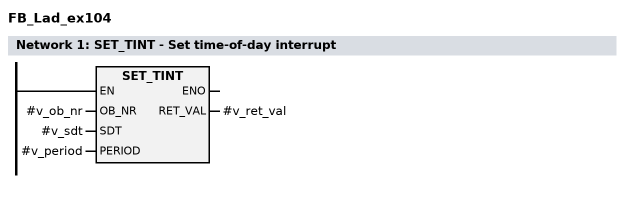
   #v_ret_val := SET_TINT(OB_NR := #v_ob_nr, SDT := #v_sdt, PERIOD := #v_period);
END_REGION
END_FUNCTION_BLOCK

FUNCTION_BLOCK "FB_Lad_ex105"   // FB30, LAD
{ S7_Optimized_Access := 'TRUE' }
   VAR_INPUT
      v_ob_nr : OB_Tod;
      v_sdt : DTL;
      v_local : Bool;
      v_period : Word;
      v_activate : Bool;
      v_ret_val : Int;
   END_VAR
BEGIN

REGION Network 1: SET_TINTL - Set time-of-day interrupt
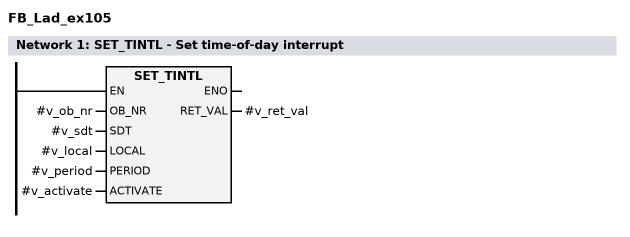
   #v_ret_val := SET_TINTL(OB_NR := #v_ob_nr,
                           SDT := #v_sdt,
                           LOCAL := #v_local,
                           PERIOD := #v_period,
                           ACTIVATE := #v_activate);
END_REGION
END_FUNCTION_BLOCK

FUNCTION_BLOCK "FB_Lad_ex106"   // FB31, LAD
{ S7_Optimized_Access := 'TRUE' }
   VAR_INPUT
      v_ob_nr : OB_Tod;
      v_ret_val : Int;
   END_VAR
BEGIN

REGION Network 1: CAN_TINT - Cancel time-of-day interrupt
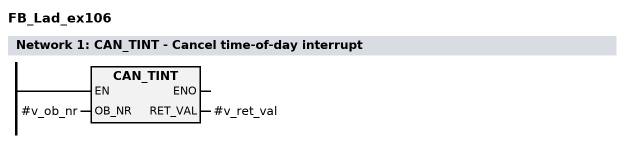
   #v_ret_val := CAN_TINT(OB_NR := #v_ob_nr);
END_REGION
END_FUNCTION_BLOCK

FUNCTION_BLOCK "FB_Lad_ex107"   // FB32, LAD
{ S7_Optimized_Access := 'TRUE' }
   VAR_INPUT
      v_ob_nr : OB_Tod;
      v_ret_val : Int;
   END_VAR
BEGIN

REGION Network 1: ACT_TINT - Enable time-of-day interrupt
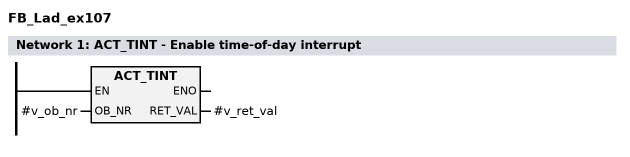
   #v_ret_val := ACT_TINT(OB_NR := #v_ob_nr);
END_REGION
END_FUNCTION_BLOCK

FUNCTION_BLOCK "FB_Lad_ex108"   // FB33, LAD
{ S7_Optimized_Access := 'TRUE' }
   VAR_INPUT
      v_ob_nr : OB_Tod;
      v_ret_val : Int;
   END_VAR
   VAR_OUTPUT
      v_status : Word;
   END_VAR
BEGIN

REGION Network 1: QRY_TINT - Query status of time-of-day interrupt
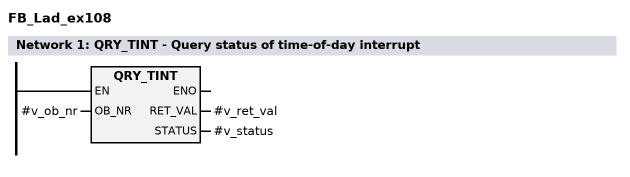
   #v_ret_val := QRY_TINT(OB_NR := #v_ob_nr, STATUS => #v_status);
END_REGION
END_FUNCTION_BLOCK

FUNCTION_BLOCK "FB_Lad_ex109"   // FB34, LAD
{ S7_Optimized_Access := 'TRUE' }
   VAR_INPUT
      v_ob_nr : Int;
      v_dtime : Time;
      v_sign : Word;
      v_ret_val : Int;
   END_VAR
BEGIN

REGION Network 1: SRT_DINT - Start time-delay interrupt
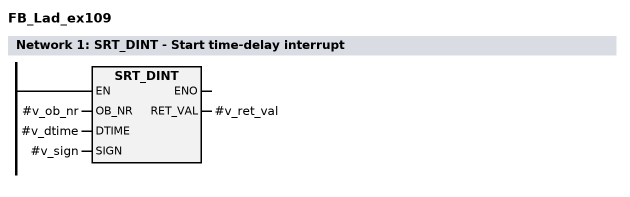
   #v_ret_val := SRT_DINT(OB_NR := #v_ob_nr, DTIME := #v_dtime, SIGN := #v_sign);
END_REGION
END_FUNCTION_BLOCK

FUNCTION_BLOCK "FB_Lad_ex110"   // FB35, LAD
{ S7_Optimized_Access := 'TRUE' }
   VAR_INPUT
      v_ob_nr : Int;
      v_ret_val : Int;
   END_VAR
BEGIN

REGION Network 1: CAN_DINT - Cancel time-delay interrupt
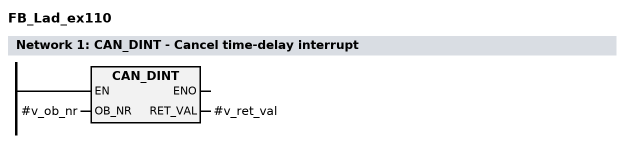
   #v_ret_val := CAN_DINT(OB_NR := #v_ob_nr);
END_REGION
END_FUNCTION_BLOCK

FUNCTION_BLOCK "FB_Lad_ex111"   // FB36, LAD
{ S7_Optimized_Access := 'TRUE' }
   VAR_INPUT
      v_ob_nr : Int;
      v_ret_val : Int;
   END_VAR
   VAR_OUTPUT
      v_status : Word;
   END_VAR
BEGIN

REGION Network 1: QRY_DINT - Query time-delay interrupt status
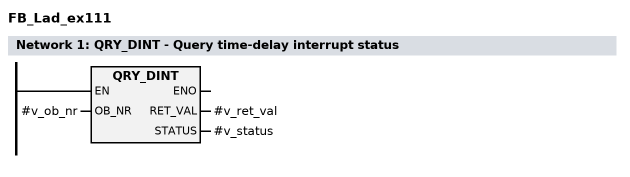
   #v_ret_val := QRY_DINT(OB_NR := #v_ob_nr, STATUS => #v_status);
END_REGION
END_FUNCTION_BLOCK

FUNCTION_BLOCK "FB_Lad_ex112"   // FB37, LAD
{ S7_Optimized_Access := 'TRUE' }
   VAR_INPUT
      v_prgflt_set_mask : DWord;
      v_accflt_set_mask : DWord;
      v_ret_val : Int;
   END_VAR
   VAR_OUTPUT
      v_prgflt_masked : DWord;
      v_accflt_masked : DWord;
   END_VAR
BEGIN

REGION Network 1: MSK_FLT - Mask synchronous error events
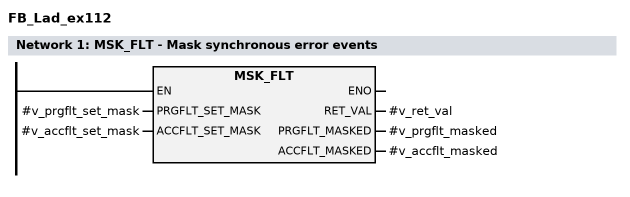
   #v_ret_val := MSK_FLT(PRGFLT_SET_MASK := #v_prgflt_set_mask,
                         ACCFLT_SET_MASK := #v_accflt_set_mask,
                         PRGFLT_MASKED => #v_prgflt_masked,
                         ACCFLT_MASKED => #v_accflt_masked);
END_REGION
END_FUNCTION_BLOCK

FUNCTION_BLOCK "FB_Lad_ex113"   // FB38, LAD
{ S7_Optimized_Access := 'TRUE' }
   VAR_INPUT
      v_prgflt_reset_mask : DWord;
      v_accflt_reset_mask : DWord;
      v_ret_val : Int;
   END_VAR
   VAR_OUTPUT
      v_prgflt_masked : DWord;
      v_accflt_masked : DWord;
   END_VAR
BEGIN

REGION Network 1: DMSK_FLT - Unmask synchronous error events
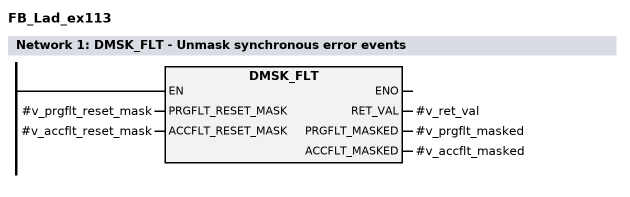
   #v_ret_val := DMSK_FLT(PRGFLT_RESET_MASK := #v_prgflt_reset_mask,
                          ACCFLT_RESET_MASK := #v_accflt_reset_mask,
                          PRGFLT_MASKED => #v_prgflt_masked,
                          ACCFLT_MASKED => #v_accflt_masked);
END_REGION
END_FUNCTION_BLOCK

FUNCTION_BLOCK "FB_Lad_ex114"   // FB39, LAD
{ S7_Optimized_Access := 'TRUE' }
   VAR_INPUT
      v_prgflt_query : DWord;
      v_accflt_query : DWord;
      v_ret_val : Int;
   END_VAR
   VAR_OUTPUT
      v_prgflt_clr : DWord;
      v_accflt_clr : DWord;
   END_VAR
BEGIN

REGION Network 1: READ_ERR - Read out event status register
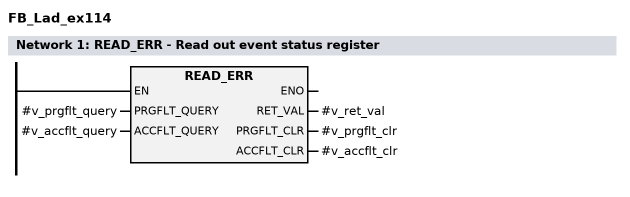
   #v_ret_val := READ_ERR(PRGFLT_QUERY := #v_prgflt_query,
                          ACCFLT_QUERY := #v_accflt_query,
                          PRGFLT_CLR => #v_prgflt_clr,
                          ACCFLT_CLR => #v_accflt_clr);
END_REGION
END_FUNCTION_BLOCK

FUNCTION_BLOCK "FB_Lad_ex115"   // FB40, LAD
{ S7_Optimized_Access := 'TRUE' }
   VAR_INPUT
      v_mode : Byte;
      v_ob_nr : Int;
      v_ret_val : Int;
   END_VAR
BEGIN

REGION Network 1: DIS_IRT - Disable interrupt event
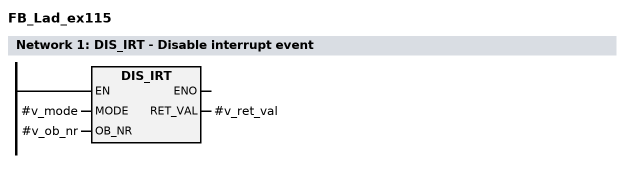
   #v_ret_val := DIS_IRT(MODE := #v_mode, OB_NR := #v_ob_nr);
END_REGION
END_FUNCTION_BLOCK

FUNCTION_BLOCK "FB_Lad_ex116"   // FB41, LAD
{ S7_Optimized_Access := 'TRUE' }
   VAR_INPUT
      v_mode : Byte;
      v_ob_nr : Int;
      v_ret_val : Int;
   END_VAR
BEGIN

REGION Network 1: EN_IRT - Enable interrupt event
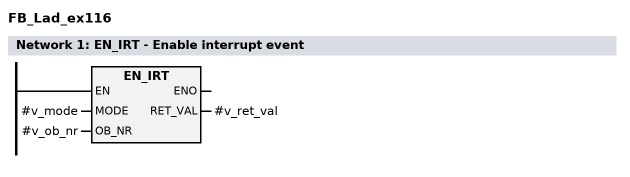
   #v_ret_val := EN_IRT(MODE := #v_mode, OB_NR := #v_ob_nr);
END_REGION
END_FUNCTION_BLOCK

FUNCTION_BLOCK "FB_Lad_ex117"   // FB42, LAD
{ S7_Optimized_Access := 'TRUE' }
   VAR_INPUT
      v_ret_val : Int;
   END_VAR
BEGIN

REGION Network 1: DIS_AIRT - Delay execution of higher priority interrupts and asynchronous error events
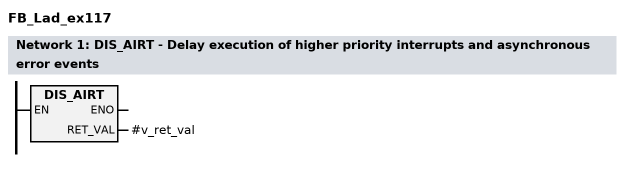
   #v_ret_val := DIS_AIRT();
END_REGION
END_FUNCTION_BLOCK

FUNCTION_BLOCK "FB_Lad_ex118"   // FB43, LAD
{ S7_Optimized_Access := 'TRUE' }
   VAR_INPUT
      v_ret_val : Int;
   END_VAR
BEGIN

REGION Network 1: EN_AIRT - Enable execution of higher priority interrupts and asynchronous error events
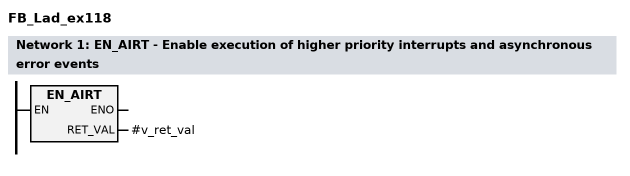
   #v_ret_val := EN_AIRT();
END_REGION
END_FUNCTION_BLOCK

FUNCTION_BLOCK "FB_Lad_ex120"   // FB44, LAD
{ S7_Optimized_Access := 'TRUE' }
   VAR_INPUT
      v_alarm : ALARM_BASE;
   END_VAR
   VAR_OUTPUT
      v_alarmstate : Byte;
      v_error : Bool;
      v_status : Word;
   END_VAR
BEGIN

REGION Network 1: Get_AlarmState - Output alarm status
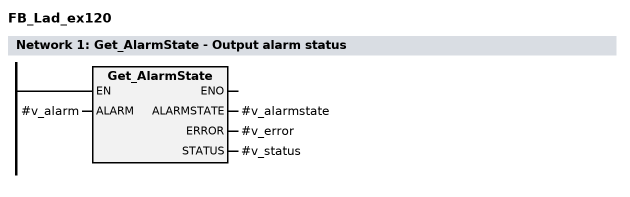
   // no SCL statement known for Get_AlarmState: written as a call
   Get_AlarmState(Alarm := #v_alarm, AlarmState => #v_alarmstate, Error => #v_error, STATUS => #v_status);
END_REGION
END_FUNCTION_BLOCK

FUNCTION_BLOCK "FB_Lad_ex121"   // FB45, LAD
{ S7_Optimized_Access := 'TRUE' }
   VAR_INPUT
      v_mode : UInt;
      v_textid : UInt;
      v_textlistid : UInt;
      v_ret_val : Int;
   END_VAR
   VAR_IN_OUT
      v_assocvalues : AssocValues;
   END_VAR
BEGIN

REGION Network 1: Gen_UsrMsg - Generate user diagnostic alarms
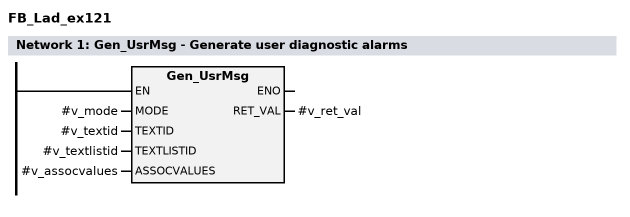
   // no SCL statement known for Gen_UsrMsg: written as a call
   #v_ret_val := Gen_UsrMsg(Mode := #v_mode,
                           TextID := #v_textid,
                           TextListID := #v_textlistid,
                           AssocValues := #v_assocvalues);
END_REGION
END_FUNCTION_BLOCK

FUNCTION_BLOCK "FB_Lad_ex123"   // FB46, LAD
{ S7_Optimized_Access := 'TRUE' }
   VAR_INPUT
      v_mode : UInt;
   END_VAR
   VAR_OUTPUT
      v_error : Bool;
      v_status : Word;
   END_VAR
BEGIN

REGION Network 1: Ack_Alarms - Acknowledge alarms
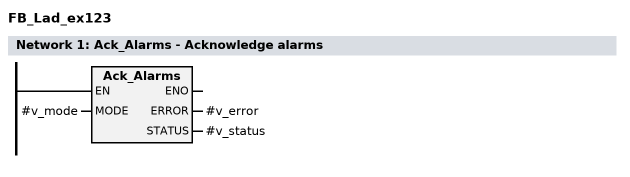
   // no SCL statement known for Ack_Alarms: written as a call
   Ack_Alarms(MODE := #v_mode, ERROR => #v_error, STATUS => #v_status);
END_REGION
END_FUNCTION_BLOCK

FUNCTION_BLOCK "FB_Lad_ex125"   // FB47, LAD
{ S7_Optimized_Access := 'TRUE' }
   VAR_INPUT
      v_mode : UInt;
      v_ob : OB_Any;
      v_ret_val : Int;
   END_VAR
   VAR_IN_OUT
      v_info : Variant;
   END_VAR
BEGIN

REGION Network 1: RT_INFO - Read out runtime statistics
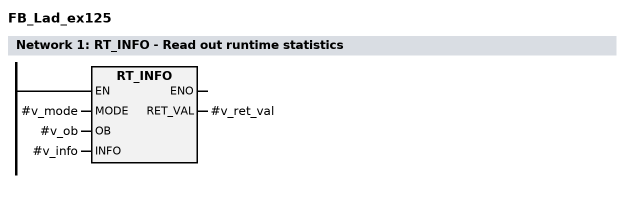
   #v_ret_val := RT_INFO(MODE := #v_mode, OB := #v_ob, INFO := #v_info);
END_REGION
END_FUNCTION_BLOCK

FUNCTION_BLOCK "FB_Lad_ex126"   // FB48, LAD
{ S7_Optimized_Access := 'TRUE' }
   VAR_INPUT
      v_laddr : Hw_Io;
      v_led : UInt;
      v_ret_val : Int;
   END_VAR
BEGIN

REGION Network 1: LED - Read LED status
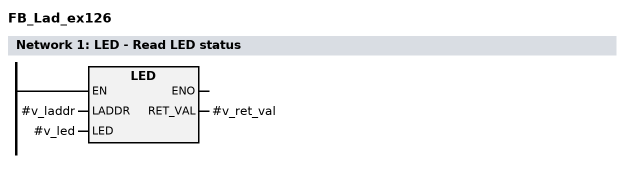
   #v_ret_val := LED(LADDR := #v_laddr, LED := #v_led);
END_REGION
END_FUNCTION_BLOCK

FUNCTION_BLOCK "FB_Lad_ex130"   // FB49, LAD
{ S7_Optimized_Access := 'TRUE' }
   VAR_INPUT
      v_laddr : Hw_IoSystem;
      v_mode : UInt;
      v_ret_val : Int;
   END_VAR
   VAR_IN_OUT
      v_state : Variant;
   END_VAR
BEGIN

REGION Network 1: DeviceStates - Read module status information in an IO system
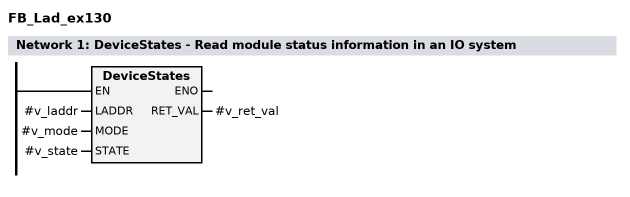
   // no SCL statement known for DeviceStates: written as a call
   #v_ret_val := DeviceStates(LADDR := #v_laddr, MODE := #v_mode, STATE := #v_state);
END_REGION
END_FUNCTION_BLOCK

FUNCTION_BLOCK "FB_Lad_ex131"   // FB50, LAD
{ S7_Optimized_Access := 'TRUE' }
   VAR_INPUT
      v_laddr : Hw_Device;
      v_mode : UInt;
      v_ret_val : Int;
   END_VAR
   VAR_IN_OUT
      v_state : Variant;
   END_VAR
BEGIN

REGION Network 1: ModuleStates - Read module status information of a module
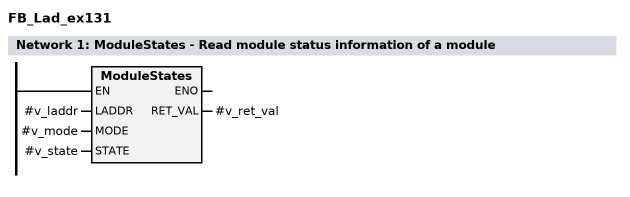
   // no SCL statement known for ModuleStates: written as a call
   #v_ret_val := ModuleStates(LADDR := #v_laddr, MODE := #v_mode, STATE := #v_state);
END_REGION
END_FUNCTION_BLOCK

FUNCTION_BLOCK "FB_Lad_ex132"   // FB51, LAD
{ S7_Optimized_Access := 'TRUE' }
   VAR_INPUT
      v_laddr : Hw_Any;
      v_mode : UInt;
      v_ret_val : Int;
   END_VAR
   VAR_IN_OUT
      v_diagevent : DiagnosticDetail;
   END_VAR
BEGIN

REGION Network 1: GEN_DIAG - Generate diagnostics information
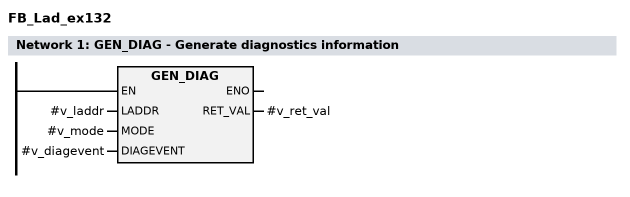
   #v_ret_val := GEN_DIAG(LADDR := #v_laddr, MODE := #v_mode, DiagEvent := #v_diagevent);
END_REGION
END_FUNCTION_BLOCK

FUNCTION_BLOCK "FB_Lad_ex133"   // FB52, LAD
{ S7_Optimized_Access := 'TRUE' }
   VAR_INPUT
      v_mode : UInt;
      v_laddr : Hw_Any;
      v_ret_val : Int;
   END_VAR
   VAR_OUTPUT
      v_cnt_diag : UInt;
   END_VAR
   VAR_IN_OUT
      v_diag : Variant;
      v_detail : Variant;
   END_VAR
BEGIN

REGION Network 1: GET_DIAG - Read diagnostic information
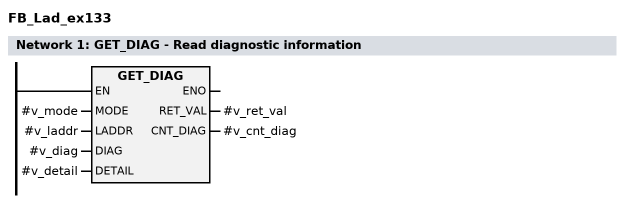
   #v_ret_val := GET_DIAG(MODE := #v_mode,
                          LADDR := #v_laddr,
                          DIAG := #v_diag,
                          DETAIL := #v_detail,
                          CNT_DIAG => #v_cnt_diag);
END_REGION
END_FUNCTION_BLOCK

FUNCTION_BLOCK "FB_Lad_ex147"   // FB53, LAD
{ S7_Optimized_Access := 'TRUE' }
   VAR_INPUT
      v_req : Bool;
      v_low_limit : UInt;
      v_up_limit : UInt;
      v_count : UDInt;
      v_attrib : Byte;
      v_srcblk : Variant;
      v_ret_val : Int;
   END_VAR
   VAR_OUTPUT
      v_busy : Bool;
      v_db_num : UInt;
   END_VAR
BEGIN

REGION Network 1: CREATE_DB - Create data block
